{attribute 'qualified_only'}
{attribute 'strict'}
{attribute 'to_string'}
TYPE E_PickStep :
(
    Undefined      := 0,
    Idle           := 10,
    LowerToPick    := 20,
    Grip           := 30,
    RaiseWithPart  := 40,
    SlideOut       := 50,
    LowerToPlace   := 60,
    ClampPart      := 65,
    OpenGripper    := 70,
    RaiseEmpty     := 80,
    ReleaseFixture := 85,
    SlideIn        := 90,
    Done           := 100,
    Error          := 900
);
END_TYPE

(* stored: Version 1.1.0.1
   DUT E_PickStep: Id {39db470c-0406-495a-9b1f-6816643f086f} *)
